INTERFACE I_Ups EXTENDS I_Module

METHOD M_Cycle
END_METHOD

PROPERTY UpsState : ST_UpsState
GET
END_GET
END_PROPERTY

METHOD M_RequestCommand : BOOL
VAR_INPUT i_eCommand : E_UpsCommand; END_VAR
END_METHOD

METHOD M_SetParameter : BOOL
VAR_INPUT i_nAddress : WORD; i_wRawValue : WORD; END_VAR
END_METHOD

END_INTERFACE

(* stored: Version 1.1.0.1, ProductVersion 3.1.4024.15
   Itf I_Ups: Id {8028375b-48c3-463b-a841-70073e1cf4d9}
   Method M_Cycle: Id {8a964840-86b8-4bac-85dd-b74edcd1c425}
   Property UpsState: Id {663c5d05-48c4-4a40-ba83-ad012582bd9c}
   Get Get: Id {a3a5fb98-8f91-42ac-ac07-5a846eb7f40c}
   Method M_RequestCommand: Id {4e32ad59-8a82-4f4a-9a4c-dc890aa4708e}
   Method M_SetParameter: Id {a7fe4f11-b251-4301-a30b-f73824f11b9d} *)
